(* IEC 61131-3 sources: codesys-ai-industrial-robot-control/plc/src/Interfaces/I_AlarmSink, 3 files *)

(* ---- Clear.st ---- *)
// The alarm condition has gone; the alarm stays listed until acknowledged.
METHOD Clear
VAR_INPUT
    eId : E_AlarmId;
END_VAR

(* ---- Raise.st ---- *)
// Raise an alarm; raising an already active alarm has no effect.
METHOD Raise
VAR_INPUT
    eId : E_AlarmId;
END_VAR

(* ---- RaiseEvent.st ---- *)
// One-shot event (no lasting condition): listed unacknowledged, never active; raised again on
// every occurrence.
METHOD RaiseEvent
VAR_INPUT
    eId : E_AlarmId;
END_VAR
